// LS Electric XG5000 project: PLC MMI 2026 SCADA PLC 1
// PLC LSPLC
// module base 0 slot 0: Input/Output Module:XBC-DR64H (DC 24V Input, Relay Output, 64 Contacts)
// module base 0 slot 1: Cnet:XBL-C21A (Cnet Module(RS-232C))
// module base 0 slot 2: FEnet:XBL-EMTA (Ethernet Module, Electrical Master)

PROGRAM DataIndikatorProses (task: Scan Program)

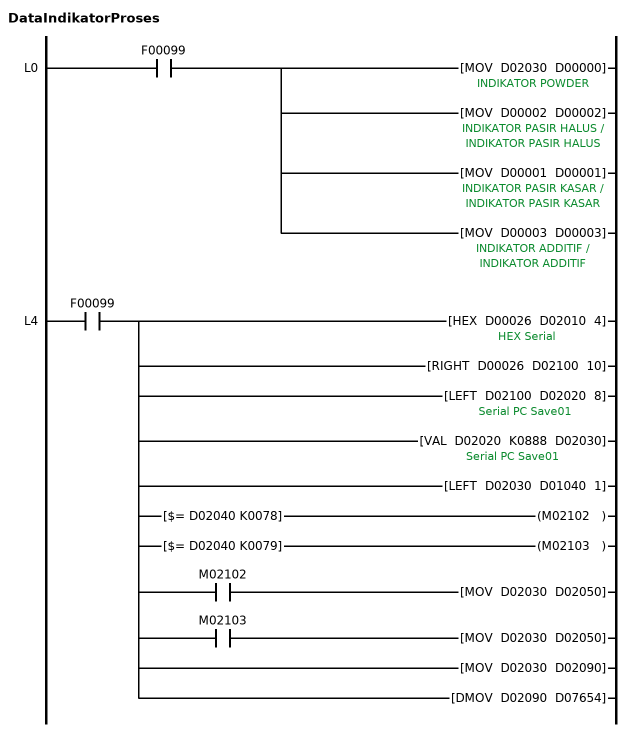
; L0
LOAD      F00099
MOV       D02030 D00000	// INDIKATOR POWDER
MOV       D00002 D00002	// INDIKATOR PASIR HALUS / INDIKATOR PASIR HALUS
MOV       D00001 D00001	// INDIKATOR PASIR KASAR / INDIKATOR PASIR KASAR
MOV       D00003 D00003	// INDIKATOR ADDITIF / INDIKATOR ADDITIF
; L4
LOAD      F00099
HEX       D00026 D02010 4	// HEX Serial
RIGHT     D00026 D02100 10
LEFT      D02100 D02020 8	// Serial PC Save01
VAL       D02020 K0888 D02030	// Serial PC Save01
LEFT      D02030 D01040 1
MPUSH
AND$=     D02040 K0078
OUT       M02102
MLOAD
AND$=     D02040 K0079
OUT       M02103
MLOAD
AND       M02102
MOV       D02030 D02050
MLOAD
AND       M02103
MOV       D02030 D02050
MPOP
MOV       D02030 D02090
DMOV      D02090 D07654

PROGRAM DataInverter (task: Scan Program)

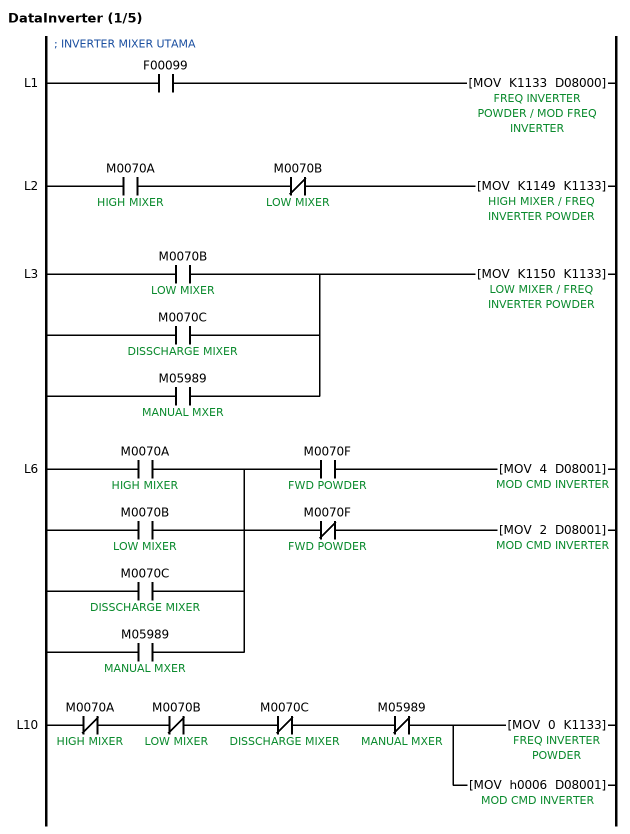
// INVERTER MIXER UTAMA
; L1
LOAD      F00099
MOV       K1133 D08000	// FREQ INVERTER POWDER / MOD FREQ INVERTER
; L2
LOAD      M0070A	// HIGH MIXER 
AND NOT   M0070B	// LOW MIXER 
MOV       K1149 K1133	// HIGH MIXER / FREQ INVERTER POWDER
; L3
LOAD      M0070B	// LOW MIXER 
OR        M0070C	// DISSCHARGE MIXER 
OR        M05989	// MANUAL MXER
MOV       K1150 K1133	// LOW MIXER / FREQ INVERTER POWDER
; L6
LOAD      M0070A	// HIGH MIXER 
OR        M0070B	// LOW MIXER 
OR        M0070C	// DISSCHARGE MIXER 
OR        M05989	// MANUAL MXER
MPUSH
AND       M0070F	// FWD POWDER
MOV       4 D08001	// MOD CMD INVERTER
MPOP
AND NOT   M0070F	// FWD POWDER
MOV       2 D08001	// MOD CMD INVERTER
; L10
LOAD NOT  M0070A	// HIGH MIXER 
AND NOT   M0070B	// LOW MIXER 
AND NOT   M0070C	// DISSCHARGE MIXER 
AND NOT   M05989	// MANUAL MXER
MOV       0 K1133	// FREQ INVERTER POWDER
MOV       h0006 D08001	// MOD CMD INVERTER

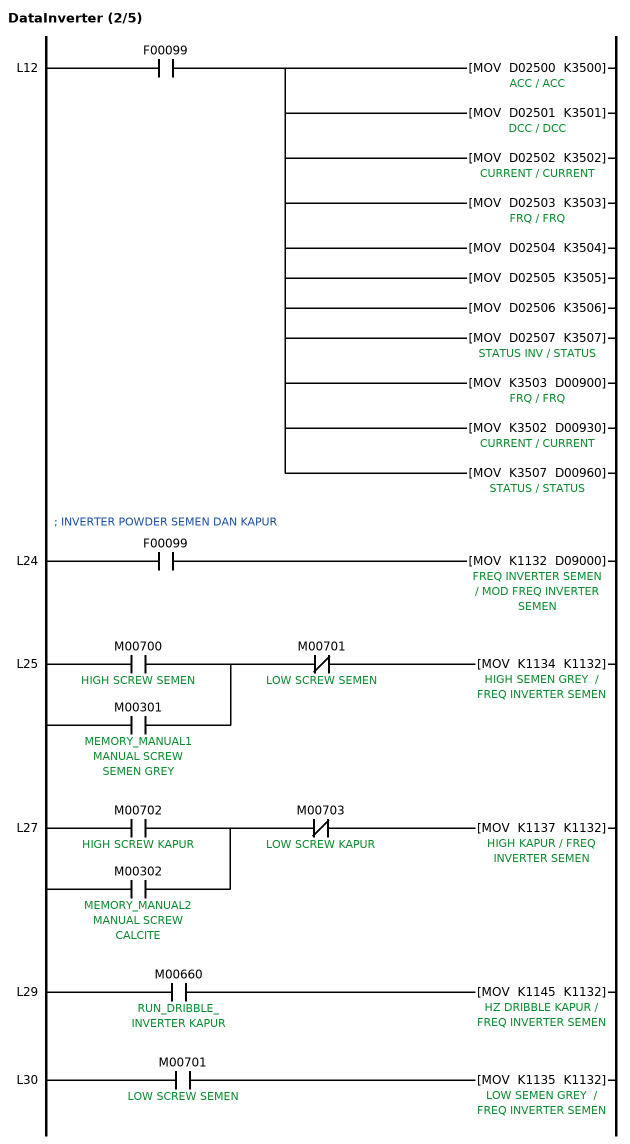
; L12
LOAD      F00099
MOV       D02500 K3500	// ACC / ACC
MOV       D02501 K3501	// DCC / DCC
MOV       D02502 K3502	// CURRENT / CURRENT
MOV       D02503 K3503	// FRQ / FRQ
MOV       D02504 K3504
MOV       D02505 K3505
MOV       D02506 K3506
MOV       D02507 K3507	// STATUS INV / STATUS
MOV       K3503 D00900	// FRQ / FRQ
MOV       K3502 D00930	// CURRENT / CURRENT
MOV       K3507 D00960	// STATUS / STATUS
// INVERTER POWDER SEMEN DAN KAPUR
; L24
LOAD      F00099
MOV       K1132 D09000	// FREQ INVERTER SEMEN  / MOD FREQ INVERTER SEMEN
; L25
LOAD      M00700	// HIGH SCREW SEMEN
OR        M00301	// MEMORY_MANUAL1 MANUAL SCREW SEMEN GREY 
AND NOT   M00701	// LOW SCREW SEMEN
MOV       K1134 K1132	// HIGH SEMEN GREY  / FREQ INVERTER SEMEN 
; L27
LOAD      M00702	// HIGH SCREW KAPUR
OR        M00302	// MEMORY_MANUAL2 MANUAL SCREW CALCITE
AND NOT   M00703	// LOW SCREW KAPUR
MOV       K1137 K1132	// HIGH KAPUR / FREQ INVERTER SEMEN 
; L29
LOAD      M00660	// RUN_DRIBBLE_INVERTER KAPUR
MOV       K1145 K1132	// HZ DRIBBLE KAPUR / FREQ INVERTER SEMEN 
; L30
LOAD      M00701	// LOW SCREW SEMEN
MOV       K1135 K1132	// LOW SEMEN GREY  / FREQ INVERTER SEMEN 

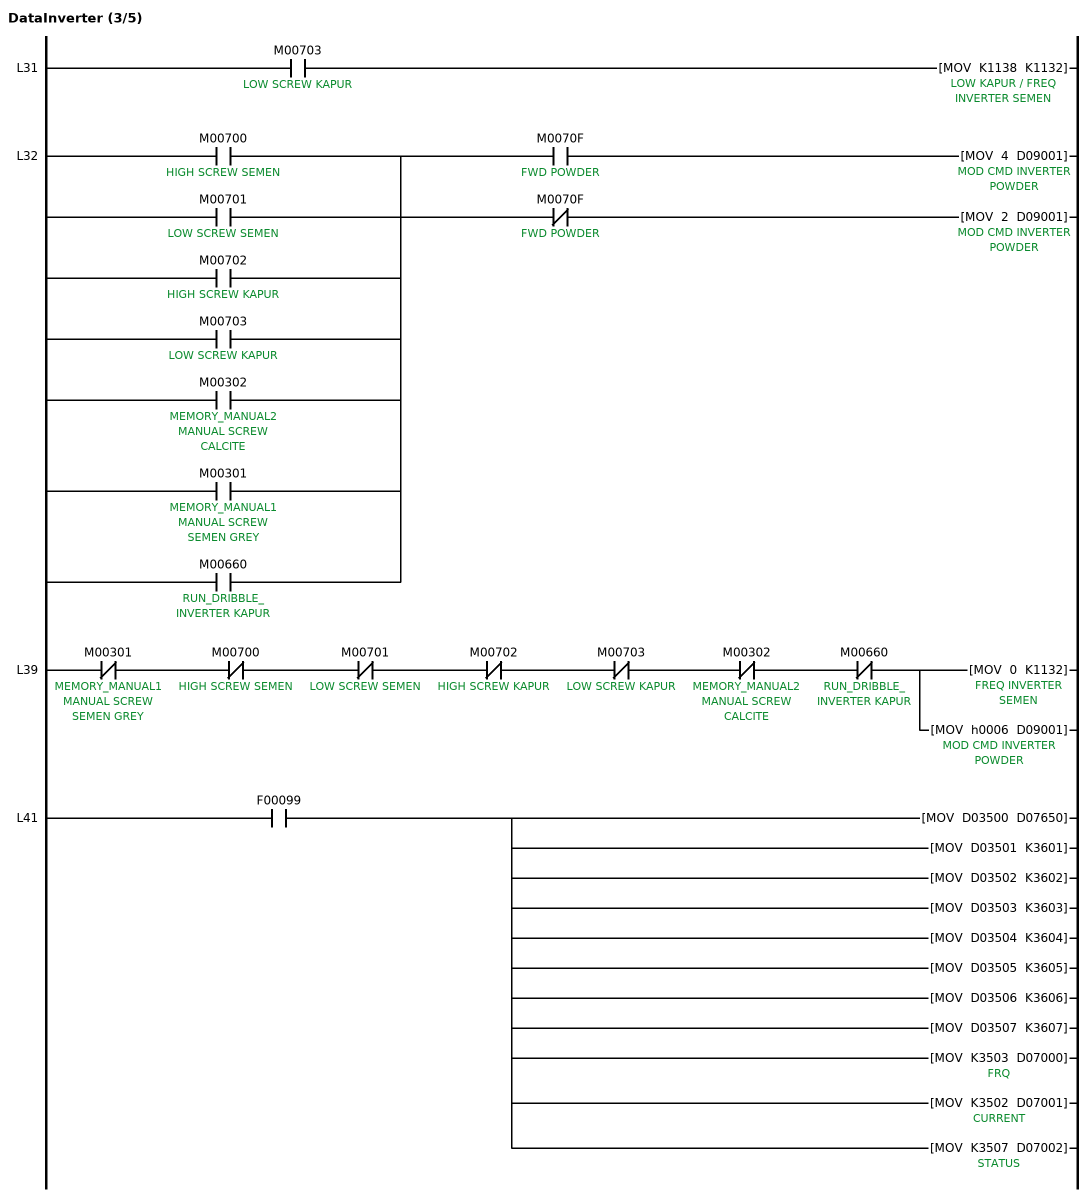
; L31
LOAD      M00703	// LOW SCREW KAPUR
MOV       K1138 K1132	// LOW KAPUR / FREQ INVERTER SEMEN 
; L32
LOAD      M00700	// HIGH SCREW SEMEN
OR        M00701	// LOW SCREW SEMEN
OR        M00702	// HIGH SCREW KAPUR
OR        M00703	// LOW SCREW KAPUR
OR        M00302	// MEMORY_MANUAL2 MANUAL SCREW CALCITE
OR        M00301	// MEMORY_MANUAL1 MANUAL SCREW SEMEN GREY 
OR        M00660	// RUN_DRIBBLE_INVERTER KAPUR
MPUSH
AND       M0070F	// FWD POWDER
MOV       4 D09001	// MOD CMD INVERTER POWDER
MPOP
AND NOT   M0070F	// FWD POWDER
MOV       2 D09001	// MOD CMD INVERTER POWDER
; L39
LOAD NOT  M00301	// MEMORY_MANUAL1 MANUAL SCREW SEMEN GREY 
AND NOT   M00700	// HIGH SCREW SEMEN
AND NOT   M00701	// LOW SCREW SEMEN
AND NOT   M00702	// HIGH SCREW KAPUR
AND NOT   M00703	// LOW SCREW KAPUR
AND NOT   M00302	// MEMORY_MANUAL2 MANUAL SCREW CALCITE
AND NOT   M00660	// RUN_DRIBBLE_INVERTER KAPUR
MOV       0 K1132	// FREQ INVERTER SEMEN 
MOV       h0006 D09001	// MOD CMD INVERTER POWDER
; L41
LOAD      F00099
MOV       D03500 D07650
MOV       D03501 K3601
MOV       D03502 K3602
MOV       D03503 K3603
MOV       D03504 K3604
MOV       D03505 K3605
MOV       D03506 K3606
MOV       D03507 K3607
MOV       K3503 D07000	// FRQ
MOV       K3502 D07001	// CURRENT
MOV       K3507 D07002	// STATUS

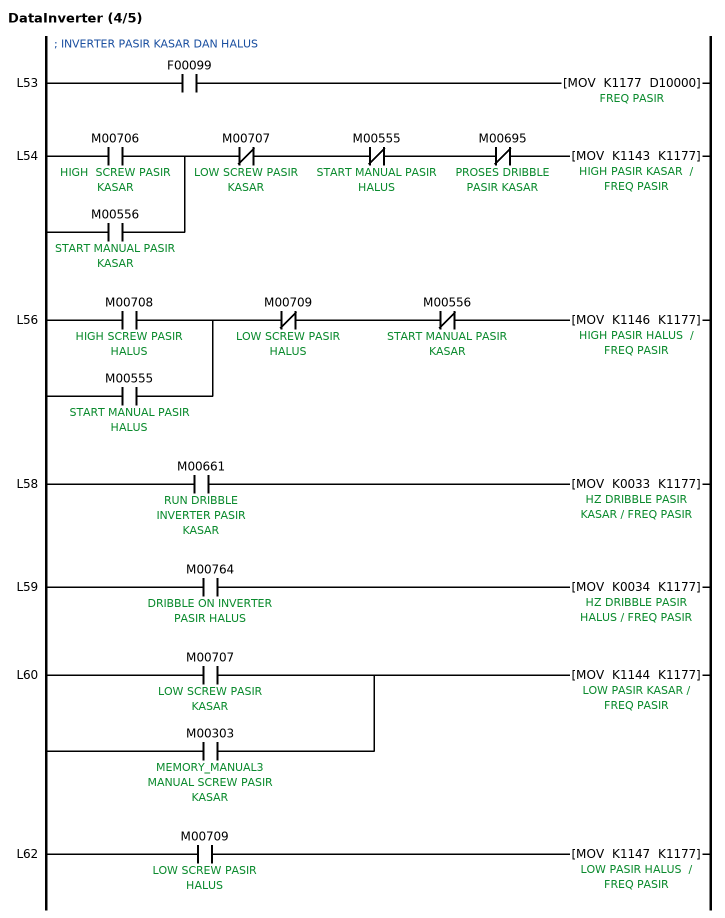
// INVERTER PASIR KASAR DAN HALUS
; L53
LOAD      F00099
MOV       K1177 D10000	// FREQ PASIR
; L54
LOAD      M00706	// HIGH  SCREW PASIR KASAR
OR        M00556	// START MANUAL PASIR KASAR
AND NOT   M00707	// LOW SCREW PASIR KASAR
AND NOT   M00555	// START MANUAL PASIR HALUS
AND NOT   M00695	// PROSES DRIBBLE PASIR KASAR
MOV       K1143 K1177	// HIGH PASIR KASAR  / FREQ PASIR
; L56
LOAD      M00708	// HIGH SCREW PASIR HALUS
OR        M00555	// START MANUAL PASIR HALUS
AND NOT   M00709	// LOW SCREW PASIR HALUS 
AND NOT   M00556	// START MANUAL PASIR KASAR
MOV       K1146 K1177	// HIGH PASIR HALUS  / FREQ PASIR
; L58
LOAD      M00661	// RUN DRIBBLE INVERTER PASIR KASAR
MOV       K0033 K1177	// HZ DRIBBLE PASIR KASAR / FREQ PASIR
; L59
LOAD      M00764	// DRIBBLE ON INVERTER PASIR HALUS
MOV       K0034 K1177	// HZ DRIBBLE PASIR HALUS / FREQ PASIR
; L60
LOAD      M00707	// LOW SCREW PASIR KASAR
OR        M00303	// MEMORY_MANUAL3 MANUAL SCREW PASIR KASAR
MOV       K1144 K1177	// LOW PASIR KASAR / FREQ PASIR
; L62
LOAD      M00709	// LOW SCREW PASIR HALUS 
MOV       K1147 K1177	// LOW PASIR HALUS  / FREQ PASIR

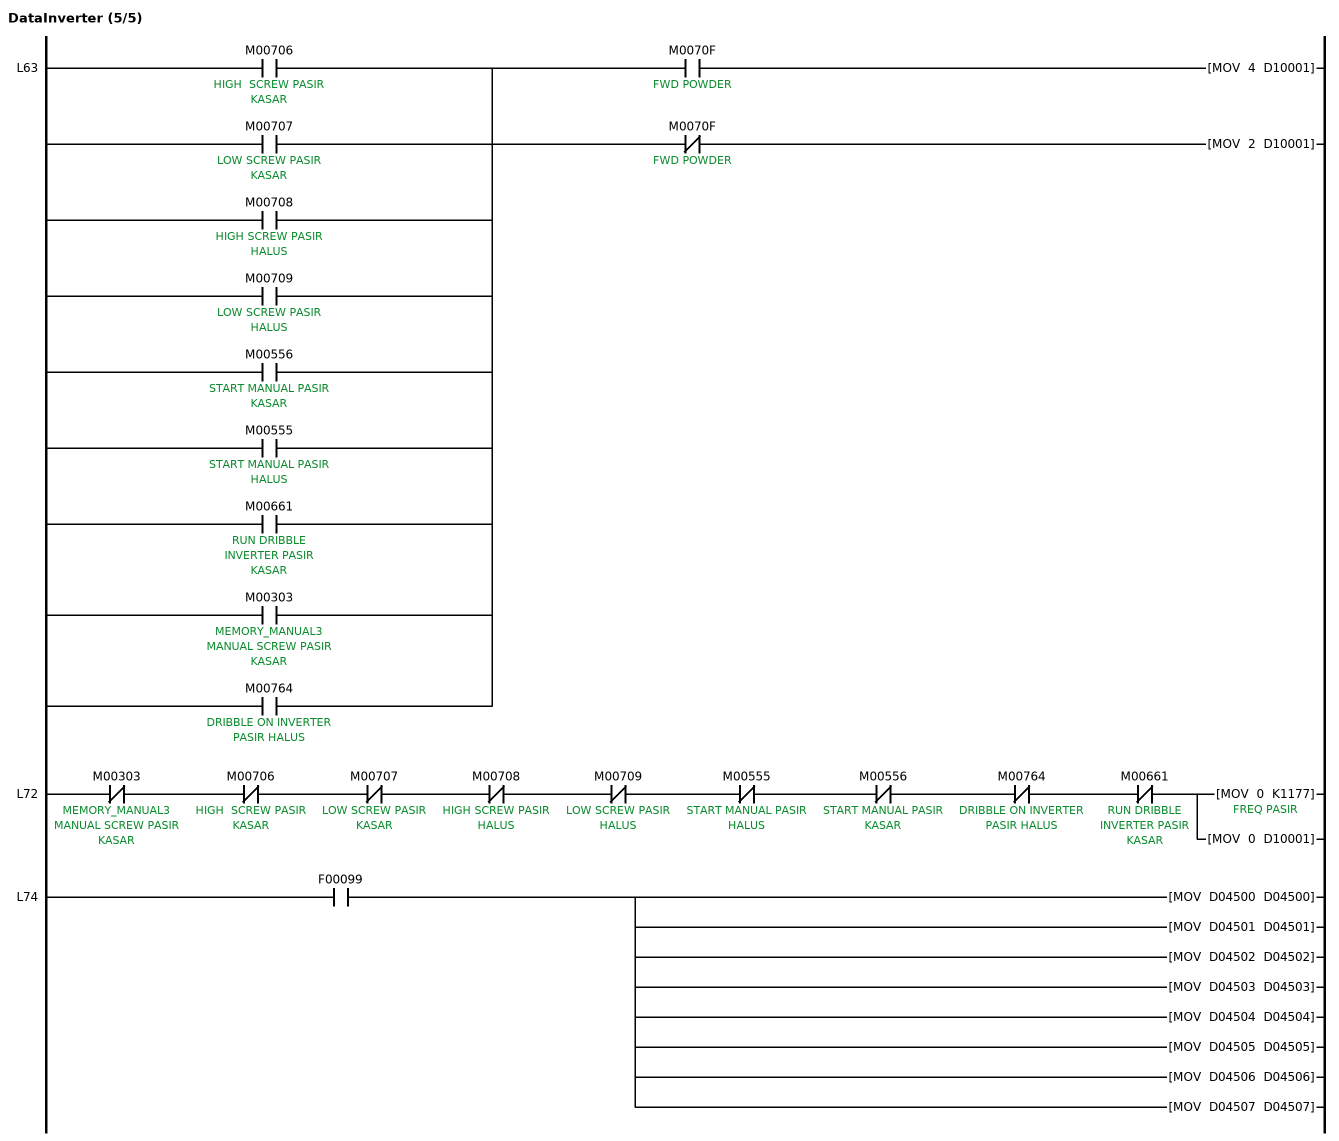
; L63
LOAD      M00706	// HIGH  SCREW PASIR KASAR
OR        M00707	// LOW SCREW PASIR KASAR
OR        M00708	// HIGH SCREW PASIR HALUS
OR        M00709	// LOW SCREW PASIR HALUS 
OR        M00556	// START MANUAL PASIR KASAR
OR        M00555	// START MANUAL PASIR HALUS
OR        M00661	// RUN DRIBBLE INVERTER PASIR KASAR
OR        M00303	// MEMORY_MANUAL3 MANUAL SCREW PASIR KASAR
OR        M00764	// DRIBBLE ON INVERTER PASIR HALUS
MPUSH
AND       M0070F	// FWD POWDER
MOV       4 D10001
MPOP
AND NOT   M0070F	// FWD POWDER
MOV       2 D10001
; L72
LOAD NOT  M00303	// MEMORY_MANUAL3 MANUAL SCREW PASIR KASAR
AND NOT   M00706	// HIGH  SCREW PASIR KASAR
AND NOT   M00707	// LOW SCREW PASIR KASAR
AND NOT   M00708	// HIGH SCREW PASIR HALUS
AND NOT   M00709	// LOW SCREW PASIR HALUS 
AND NOT   M00555	// START MANUAL PASIR HALUS
AND NOT   M00556	// START MANUAL PASIR KASAR
AND NOT   M00764	// DRIBBLE ON INVERTER PASIR HALUS
AND NOT   M00661	// RUN DRIBBLE INVERTER PASIR KASAR
MOV       0 K1177	// FREQ PASIR
MOV       0 D10001
; L74
LOAD      F00099
MOV       D04500 D04500
MOV       D04501 D04501
MOV       D04502 D04502
MOV       D04503 D04503
MOV       D04504 D04504
MOV       D04505 D04505
MOV       D04506 D04506
MOV       D04507 D04507

PROGRAM FormulaSet (task: Scan Program)

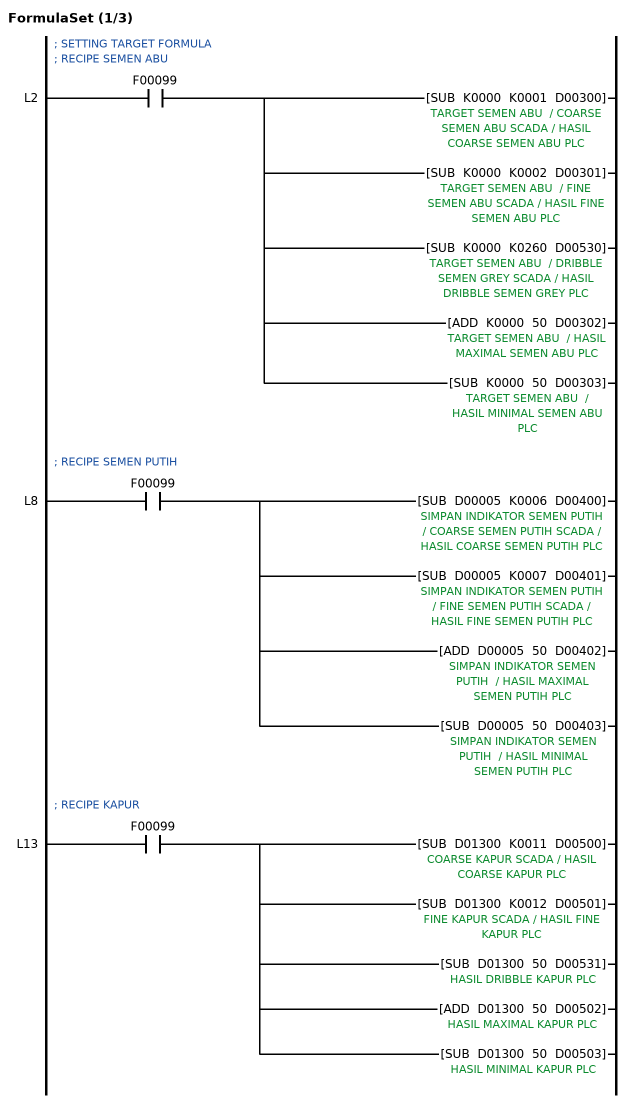
// SETTING TARGET FORMULA
// RECIPE SEMEN ABU
; L2
LOAD      F00099
SUB       K0000 K0001 D00300	// TARGET SEMEN ABU  / COARSE SEMEN ABU SCADA / HASIL COARSE SEMEN ABU PLC
SUB       K0000 K0002 D00301	// TARGET SEMEN ABU  / FINE SEMEN ABU SCADA / HASIL FINE SEMEN ABU PLC
SUB       K0000 K0260 D00530	// TARGET SEMEN ABU  / DRIBBLE SEMEN GREY SCADA / HASIL DRIBBLE SEMEN GREY PLC
ADD       K0000 50 D00302	// TARGET SEMEN ABU  / HASIL MAXIMAL SEMEN ABU PLC
SUB       K0000 50 D00303	// TARGET SEMEN ABU  / HASIL MINIMAL SEMEN ABU PLC
// RECIPE SEMEN PUTIH
; L8
LOAD      F00099
SUB       D00005 K0006 D00400	// SIMPAN INDIKATOR SEMEN PUTIH  / COARSE SEMEN PUTIH SCADA / HASIL COARSE SEMEN PUTIH PLC
SUB       D00005 K0007 D00401	// SIMPAN INDIKATOR SEMEN PUTIH  / FINE SEMEN PUTIH SCADA / HASIL FINE SEMEN PUTIH PLC 
ADD       D00005 50 D00402	// SIMPAN INDIKATOR SEMEN PUTIH  / HASIL MAXIMAL SEMEN PUTIH PLC 
SUB       D00005 50 D00403	// SIMPAN INDIKATOR SEMEN PUTIH  / HASIL MINIMAL SEMEN PUTIH PLC
// RECIPE KAPUR
; L13
LOAD      F00099
SUB       D01300 K0011 D00500	// COARSE KAPUR SCADA / HASIL COARSE KAPUR PLC
SUB       D01300 K0012 D00501	// FINE KAPUR SCADA / HASIL FINE KAPUR PLC 
SUB       D01300 50 D00531	// HASIL DRIBBLE KAPUR PLC 
ADD       D01300 50 D00502	// HASIL MAXIMAL KAPUR PLC 
SUB       D01300 50 D00503	// HASIL MINIMAL KAPUR PLC 

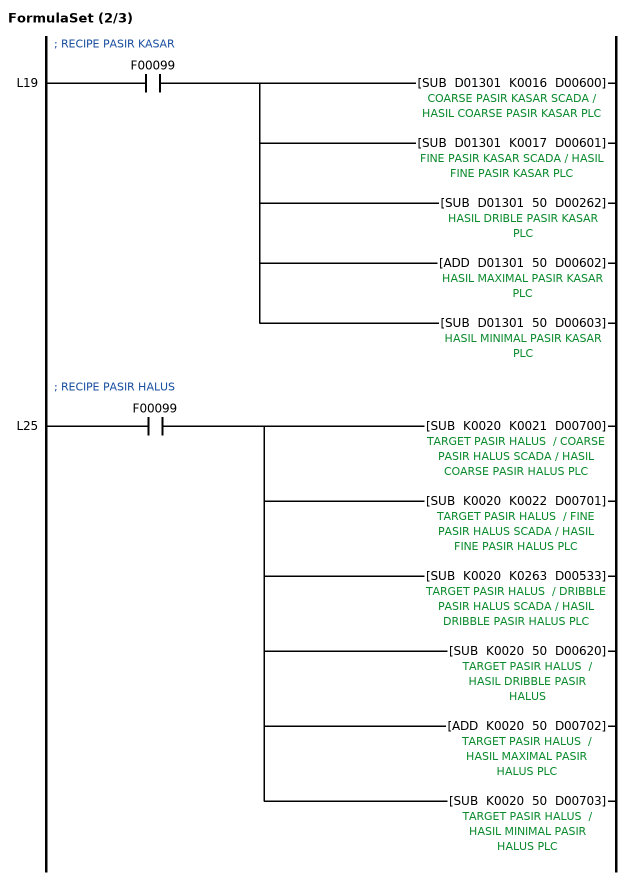
// RECIPE PASIR KASAR
; L19
LOAD      F00099
SUB       D01301 K0016 D00600	// COARSE PASIR KASAR SCADA / HASIL COARSE PASIR KASAR PLC
SUB       D01301 K0017 D00601	// FINE PASIR KASAR SCADA / HASIL FINE PASIR KASAR PLC
SUB       D01301 50 D00262	// HASIL DRIBLE PASIR KASAR PLC
ADD       D01301 50 D00602	// HASIL MAXIMAL PASIR KASAR PLC
SUB       D01301 50 D00603	// HASIL MINIMAL PASIR KASAR PLC
// RECIPE PASIR HALUS
; L25
LOAD      F00099
SUB       K0020 K0021 D00700	// TARGET PASIR HALUS  / COARSE PASIR HALUS SCADA / HASIL COARSE PASIR HALUS PLC
SUB       K0020 K0022 D00701	// TARGET PASIR HALUS  / FINE PASIR HALUS SCADA / HASIL FINE PASIR HALUS PLC
SUB       K0020 K0263 D00533	// TARGET PASIR HALUS  / DRIBBLE PASIR HALUS SCADA / HASIL DRIBBLE PASIR HALUS PLC
SUB       K0020 50 D00620	// TARGET PASIR HALUS  / HASIL DRIBBLE PASIR HALUS
ADD       K0020 50 D00702	// TARGET PASIR HALUS  / HASIL MAXIMAL PASIR HALUS PLC
SUB       K0020 50 D00703	// TARGET PASIR HALUS  / HASIL MINIMAL PASIR HALUS PLC

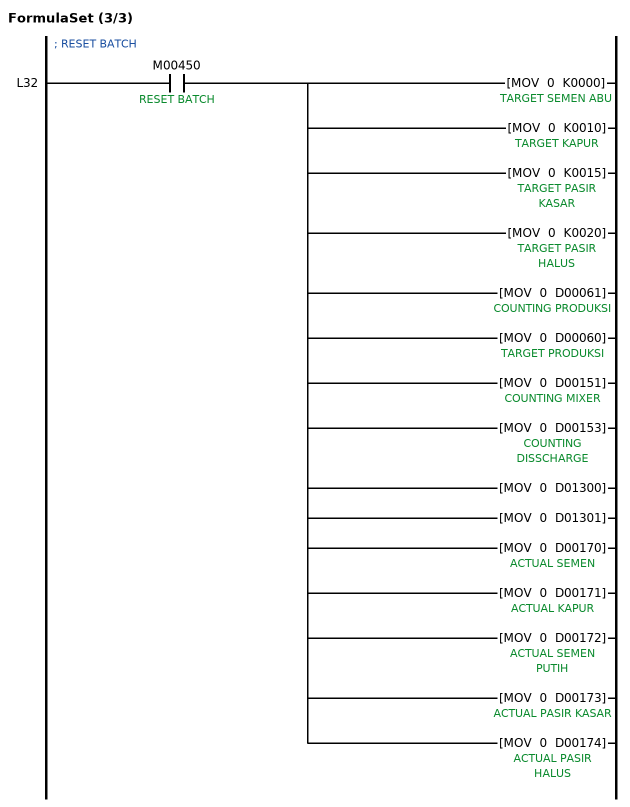
// RESET BATCH
; L32
LOAD      M00450	// RESET BATCH
MOV       0 K0000	// TARGET SEMEN ABU 
MOV       0 K0010	// TARGET KAPUR 
MOV       0 K0015	// TARGET PASIR KASAR
MOV       0 K0020	// TARGET PASIR HALUS 
MOV       0 D00061	// COUNTING PRODUKSI
MOV       0 D00060	// TARGET PRODUKSI
MOV       0 D00151	// COUNTING MIXER
MOV       0 D00153	// COUNTING DISSCHARGE
MOV       0 D01300
MOV       0 D01301
MOV       0 D00170	// ACTUAL SEMEN
MOV       0 D00171	// ACTUAL KAPUR
MOV       0 D00172	// ACTUAL SEMEN PUTIH
MOV       0 D00173	// ACTUAL PASIR KASAR
MOV       0 D00174	// ACTUAL PASIR HALUS

PROGRAM DigitalInput (task: Scan Program)

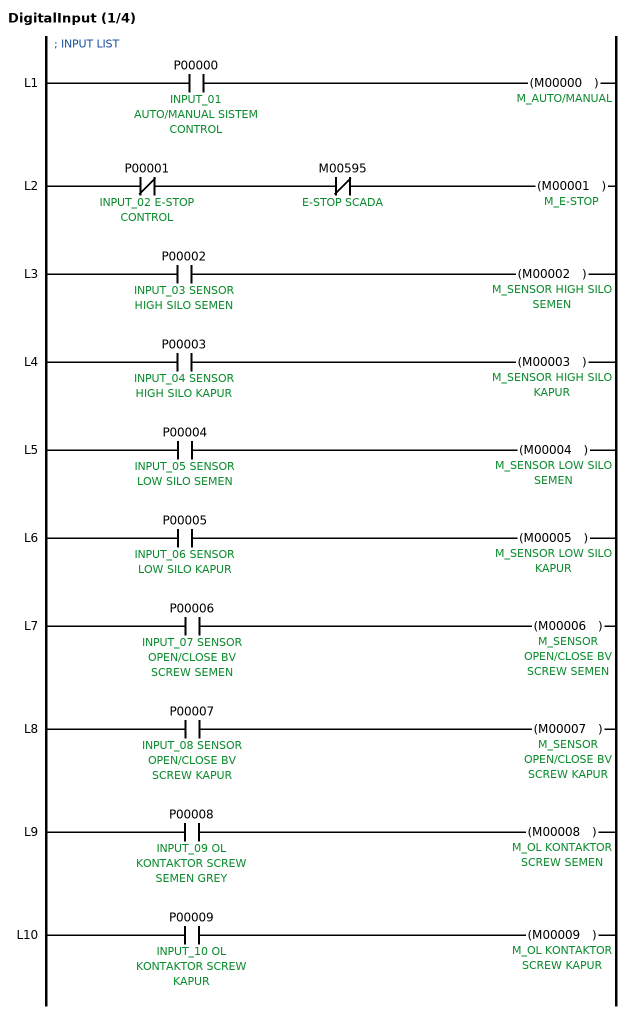
// INPUT LIST
; L1
LOAD      P00000	// INPUT_01 AUTO/MANUAL SISTEM CONTROL
OUT       M00000	// M_AUTO/MANUAL
; L2
LOAD NOT  P00001	// INPUT_02 E-STOP CONTROL 
AND NOT   M00595	// E-STOP SCADA
OUT       M00001	// M_E-STOP
; L3
LOAD      P00002	// INPUT_03 SENSOR HIGH SILO SEMEN
OUT       M00002	// M_SENSOR HIGH SILO SEMEN 
; L4
LOAD      P00003	// INPUT_04 SENSOR HIGH SILO KAPUR
OUT       M00003	// M_SENSOR HIGH SILO KAPUR
; L5
LOAD      P00004	// INPUT_05 SENSOR LOW SILO SEMEN
OUT       M00004	// M_SENSOR LOW SILO SEMEN 
; L6
LOAD      P00005	// INPUT_06 SENSOR LOW SILO KAPUR
OUT       M00005	// M_SENSOR LOW SILO KAPUR
; L7
LOAD      P00006	// INPUT_07 SENSOR OPEN/CLOSE BV SCREW SEMEN
OUT       M00006	// M_SENSOR OPEN/CLOSE BV SCREW SEMEN
; L8
LOAD      P00007	// INPUT_08 SENSOR OPEN/CLOSE BV SCREW KAPUR
OUT       M00007	// M_SENSOR OPEN/CLOSE BV SCREW KAPUR
; L9
LOAD      P00008	// INPUT_09 OL KONTAKTOR SCREW SEMEN GREY 
OUT       M00008	// M_OL KONTAKTOR SCREW SEMEN
; L10
LOAD      P00009	// INPUT_10 OL KONTAKTOR SCREW KAPUR
OUT       M00009	// M_OL KONTAKTOR SCREW KAPUR

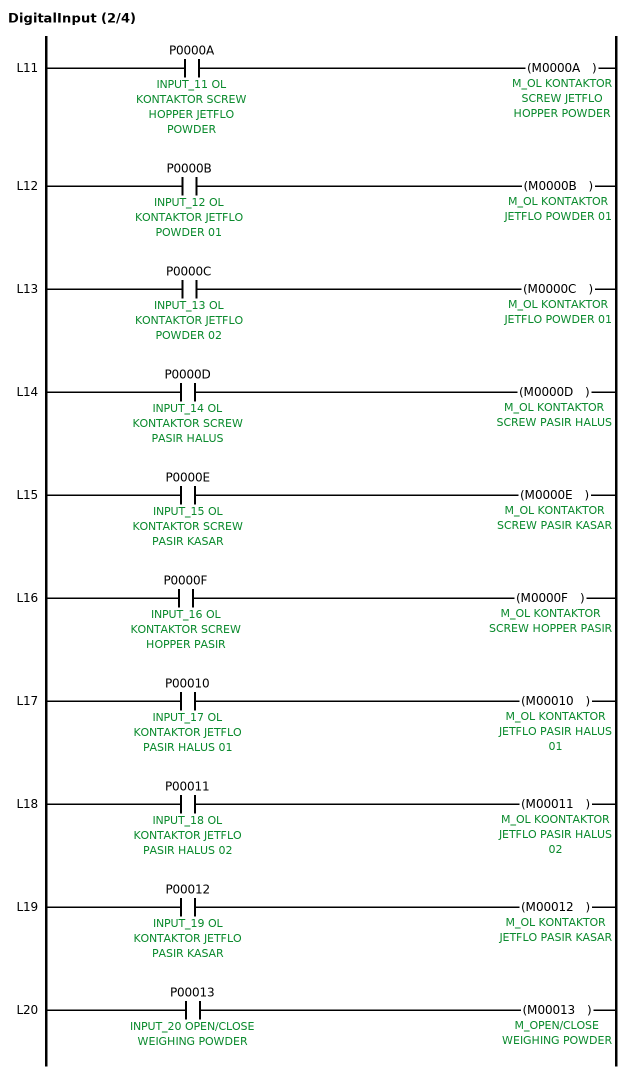
; L11
LOAD      P0000A	// INPUT_11 OL KONTAKTOR SCREW HOPPER JETFLO POWDER
OUT       M0000A	// M_OL KONTAKTOR SCREW JETFLO HOPPER POWDER
; L12
LOAD      P0000B	// INPUT_12 OL KONTAKTOR JETFLO POWDER 01
OUT       M0000B	// M_OL KONTAKTOR JETFLO POWDER 01
; L13
LOAD      P0000C	// INPUT_13 OL KONTAKTOR JETFLO POWDER 02
OUT       M0000C	// M_OL KONTAKTOR JETFLO POWDER 01
; L14
LOAD      P0000D	// INPUT_14 OL KONTAKTOR SCREW PASIR HALUS 
OUT       M0000D	// M_OL KONTAKTOR SCREW PASIR HALUS 
; L15
LOAD      P0000E	// INPUT_15 OL KONTAKTOR SCREW PASIR KASAR
OUT       M0000E	// M_OL KONTAKTOR SCREW PASIR KASAR
; L16
LOAD      P0000F	// INPUT_16 OL KONTAKTOR SCREW HOPPER PASIR 
OUT       M0000F	// M_OL KONTAKTOR SCREW HOPPER PASIR
; L17
LOAD      P00010	// INPUT_17 OL KONTAKTOR JETFLO PASIR HALUS 01
OUT       M00010	// M_OL KONTAKTOR JETFLO PASIR HALUS 01
; L18
LOAD      P00011	// INPUT_18 OL KONTAKTOR JETFLO PASIR HALUS 02
OUT       M00011	// M_OL KOONTAKTOR JETFLO PASIR HALUS 02
; L19
LOAD      P00012	// INPUT_19 OL KONTAKTOR JETFLO PASIR KASAR 
OUT       M00012	// M_OL KONTAKTOR JETFLO PASIR KASAR
; L20
LOAD      P00013	// INPUT_20 OPEN/CLOSE WEIGHING POWDER
OUT       M00013	// M_OPEN/CLOSE WEIGHING POWDER

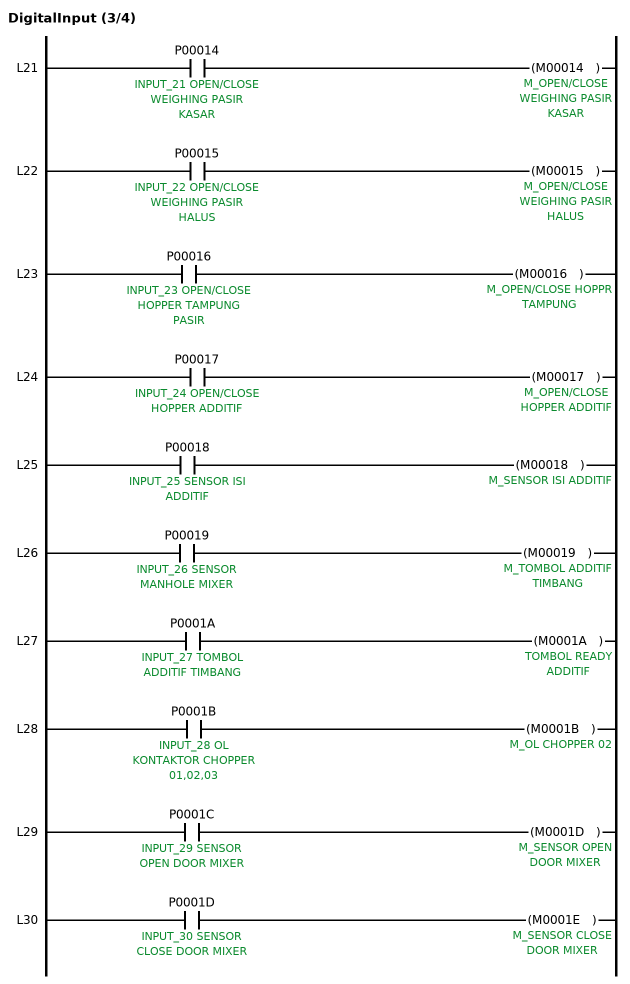
; L21
LOAD      P00014	// INPUT_21 OPEN/CLOSE WEIGHING PASIR KASAR
OUT       M00014	// M_OPEN/CLOSE WEIGHING PASIR KASAR
; L22
LOAD      P00015	// INPUT_22 OPEN/CLOSE WEIGHING PASIR HALUS
OUT       M00015	// M_OPEN/CLOSE WEIGHING PASIR HALUS 
; L23
LOAD      P00016	// INPUT_23 OPEN/CLOSE HOPPER TAMPUNG PASIR
OUT       M00016	// M_OPEN/CLOSE HOPPR TAMPUNG
; L24
LOAD      P00017	// INPUT_24 OPEN/CLOSE HOPPER ADDITIF
OUT       M00017	// M_OPEN/CLOSE HOPPER ADDITIF
; L25
LOAD      P00018	// INPUT_25 SENSOR ISI ADDITIF
OUT       M00018	// M_SENSOR ISI ADDITIF
; L26
LOAD      P00019	// INPUT_26 SENSOR MANHOLE MIXER
OUT       M00019	// M_TOMBOL ADDITIF TIMBANG
; L27
LOAD      P0001A	// INPUT_27 TOMBOL ADDITIF TIMBANG 
OUT       M0001A	// TOMBOL READY ADDITIF
; L28
LOAD      P0001B	// INPUT_28 OL KONTAKTOR CHOPPER 01,02,03
OUT       M0001B	// M_OL CHOPPER 02
; L29
LOAD      P0001C	// INPUT_29 SENSOR OPEN DOOR MIXER
OUT       M0001D	// M_SENSOR OPEN DOOR MIXER 
; L30
LOAD      P0001D	// INPUT_30 SENSOR CLOSE DOOR MIXER
OUT       M0001E	// M_SENSOR CLOSE DOOR MIXER

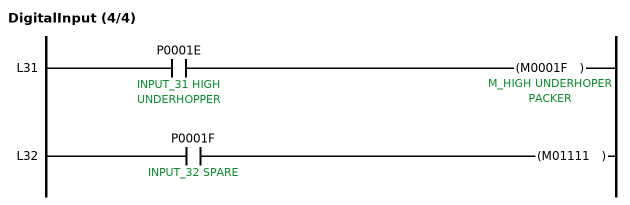
; L31
LOAD      P0001E	// INPUT_31 HIGH UNDERHOPPER
OUT       M0001F	// M_HIGH UNDERHOPER PACKER
; L32
LOAD      P0001F	// INPUT_32 SPARE
OUT       M01111

PROGRAM DigitalOutput (task: Scan Program)

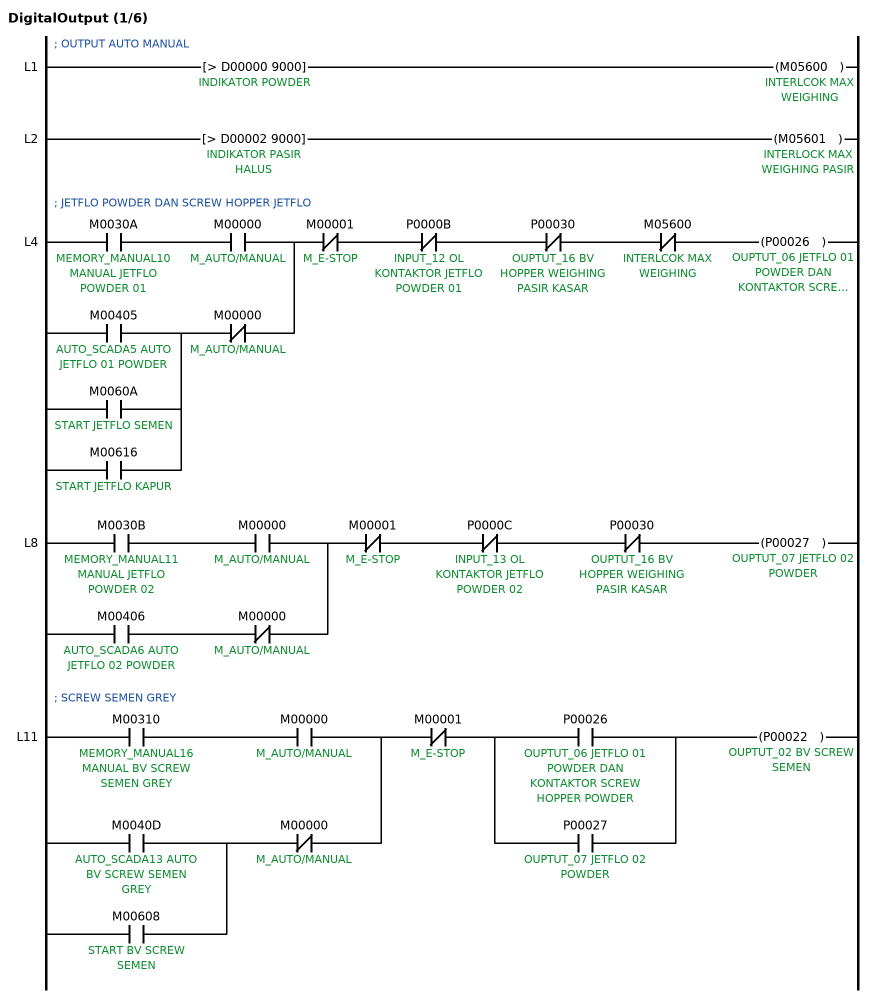
// OUTPUT AUTO MANUAL
; L1
LOAD>     D00000 9000	// INDIKATOR POWDER
OUT       M05600	// INTERLCOK MAX WEIGHING
; L2
LOAD>     D00002 9000	// INDIKATOR PASIR HALUS
OUT       M05601	// INTERLOCK MAX WEIGHING PASIR
// JETFLO POWDER DAN SCREW HOPPER JETFLO
; L4
LOAD      M0030A	// MEMORY_MANUAL10 MANUAL JETFLO POWDER 01 
AND       M00000	// M_AUTO/MANUAL
LOAD      M00405	// AUTO_SCADA5 AUTO JETFLO 01 POWDER
OR        M0060A	// START JETFLO SEMEN
OR        M00616	// START JETFLO KAPUR
AND NOT   M00000	// M_AUTO/MANUAL
OR LOAD
AND NOT   M00001	// M_E-STOP
AND NOT   P0000B	// INPUT_12 OL KONTAKTOR JETFLO POWDER 01
AND NOT   P00030	// OUPTUT_16 BV HOPPER WEIGHING PASIR KASAR
AND NOT   M05600	// INTERLCOK MAX WEIGHING
OUT       P00026	// OUPTUT_06 JETFLO 01 POWDER DAN KONTAKTOR SCREW HOPPER POWDER
; L8
LOAD      M0030B	// MEMORY_MANUAL11 MANUAL JETFLO POWDER 02 
AND       M00000	// M_AUTO/MANUAL
LOAD      M00406	// AUTO_SCADA6 AUTO JETFLO 02 POWDER
AND NOT   M00000	// M_AUTO/MANUAL
OR LOAD
AND NOT   M00001	// M_E-STOP
AND NOT   P0000C	// INPUT_13 OL KONTAKTOR JETFLO POWDER 02
AND NOT   P00030	// OUPTUT_16 BV HOPPER WEIGHING PASIR KASAR
OUT       P00027	// OUPTUT_07 JETFLO 02 POWDER 
// SCREW SEMEN GREY
; L11
LOAD      M00310	// MEMORY_MANUAL16 MANUAL BV SCREW SEMEN GREY 
AND       M00000	// M_AUTO/MANUAL
LOAD      M0040D	// AUTO_SCADA13 AUTO BV SCREW SEMEN GREY 
OR        M00608	// START BV SCREW SEMEN 
AND NOT   M00000	// M_AUTO/MANUAL
OR LOAD
AND NOT   M00001	// M_E-STOP
LOAD      P00026	// OUPTUT_06 JETFLO 01 POWDER DAN KONTAKTOR SCREW HOPPER POWDER
OR        P00027	// OUPTUT_07 JETFLO 02 POWDER 
AND LOAD
OUT       P00022	// OUPTUT_02 BV SCREW SEMEN

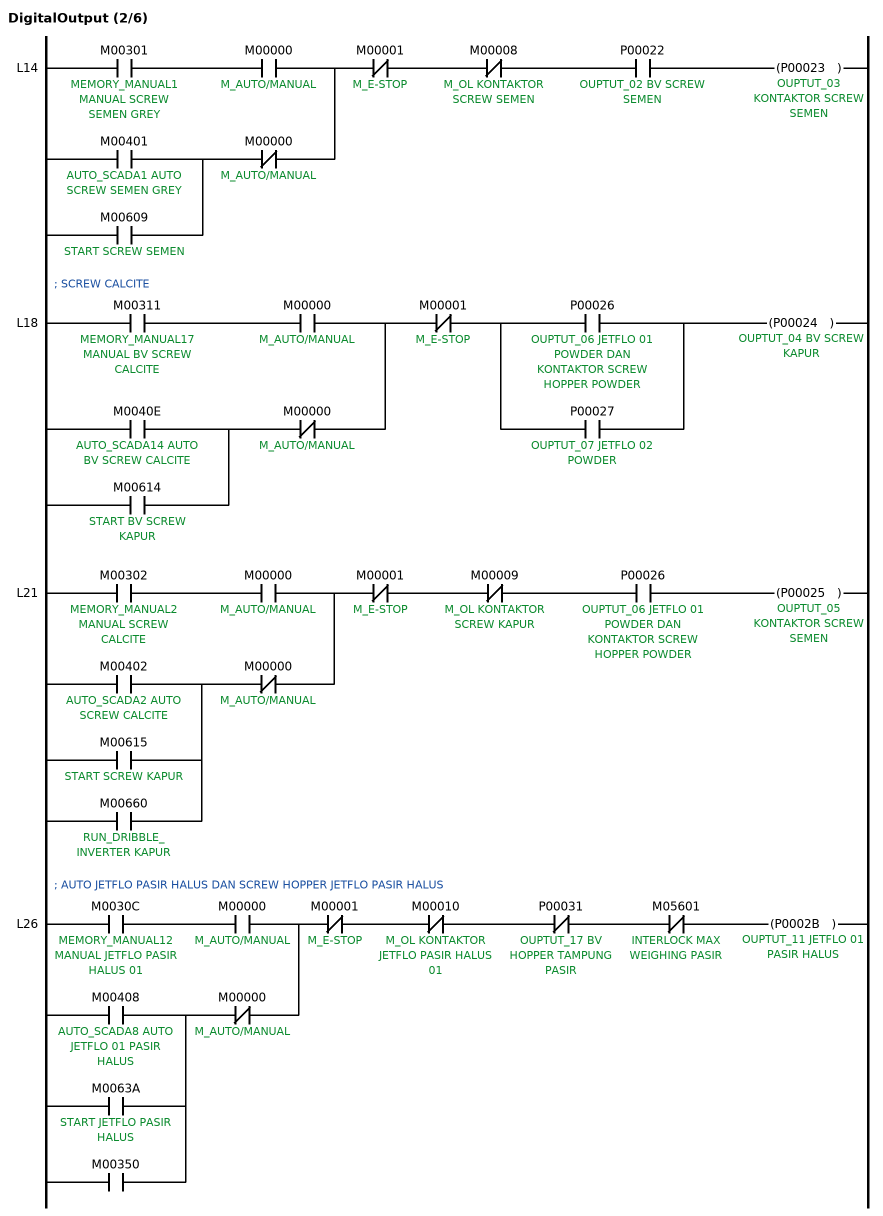
; L14
LOAD      M00301	// MEMORY_MANUAL1 MANUAL SCREW SEMEN GREY 
AND       M00000	// M_AUTO/MANUAL
LOAD      M00401	// AUTO_SCADA1 AUTO SCREW SEMEN GREY 
OR        M00609	// START SCREW SEMEN
AND NOT   M00000	// M_AUTO/MANUAL
OR LOAD
AND NOT   M00001	// M_E-STOP
AND NOT   M00008	// M_OL KONTAKTOR SCREW SEMEN
AND       P00022	// OUPTUT_02 BV SCREW SEMEN
OUT       P00023	// OUPTUT_03 KONTAKTOR SCREW SEMEN
// SCREW CALCITE
; L18
LOAD      M00311	// MEMORY_MANUAL17 MANUAL BV SCREW CALCITE
AND       M00000	// M_AUTO/MANUAL
LOAD      M0040E	// AUTO_SCADA14 AUTO BV SCREW CALCITE
OR        M00614	// START BV SCREW KAPUR
AND NOT   M00000	// M_AUTO/MANUAL
OR LOAD
AND NOT   M00001	// M_E-STOP
LOAD      P00026	// OUPTUT_06 JETFLO 01 POWDER DAN KONTAKTOR SCREW HOPPER POWDER
OR        P00027	// OUPTUT_07 JETFLO 02 POWDER 
AND LOAD
OUT       P00024	// OUPTUT_04 BV SCREW KAPUR
; L21
LOAD      M00302	// MEMORY_MANUAL2 MANUAL SCREW CALCITE
AND       M00000	// M_AUTO/MANUAL
LOAD      M00402	// AUTO_SCADA2 AUTO SCREW CALCITE
OR        M00615	// START SCREW KAPUR
OR        M00660	// RUN_DRIBBLE_INVERTER KAPUR
AND NOT   M00000	// M_AUTO/MANUAL
OR LOAD
AND NOT   M00001	// M_E-STOP
AND NOT   M00009	// M_OL KONTAKTOR SCREW KAPUR
AND       P00026	// OUPTUT_06 JETFLO 01 POWDER DAN KONTAKTOR SCREW HOPPER POWDER
OUT       P00025	// OUPTUT_05 KONTAKTOR SCREW SEMEN
// AUTO JETFLO PASIR HALUS DAN SCREW HOPPER JETFLO PASIR HALUS
; L26
LOAD      M0030C	// MEMORY_MANUAL12 MANUAL JETFLO PASIR HALUS 01 
AND       M00000	// M_AUTO/MANUAL
LOAD      M00408	// AUTO_SCADA8 AUTO JETFLO 01 PASIR HALUS 
OR        M0063A	// START JETFLO PASIR  HALUS
OR        M00350
AND NOT   M00000	// M_AUTO/MANUAL
OR LOAD
AND NOT   M00001	// M_E-STOP
AND NOT   M00010	// M_OL KONTAKTOR JETFLO PASIR HALUS 01
AND NOT   P00031	// OUPTUT_17 BV HOPPER TAMPUNG PASIR
AND NOT   M05601	// INTERLOCK MAX WEIGHING PASIR
OUT       P0002B	// OUPTUT_11 JETFLO 01 PASIR HALUS

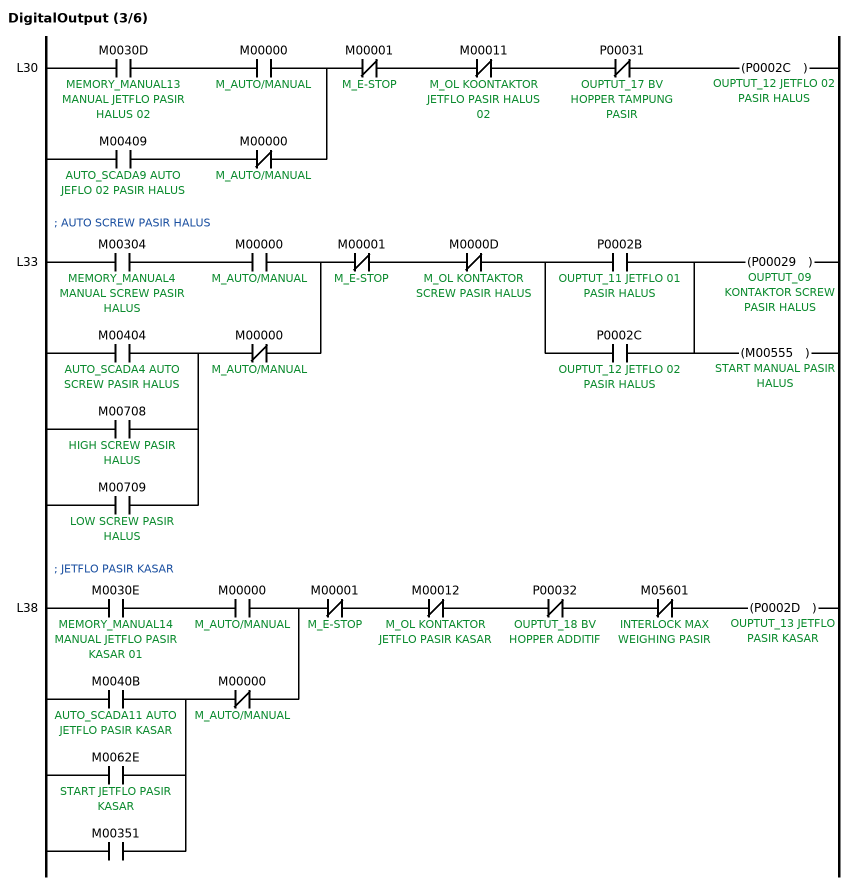
; L30
LOAD      M0030D	// MEMORY_MANUAL13 MANUAL JETFLO PASIR HALUS 02 
AND       M00000	// M_AUTO/MANUAL
LOAD      M00409	// AUTO_SCADA9 AUTO JEFLO 02 PASIR HALUS 
AND NOT   M00000	// M_AUTO/MANUAL
OR LOAD
AND NOT   M00001	// M_E-STOP
AND NOT   M00011	// M_OL KOONTAKTOR JETFLO PASIR HALUS 02
AND NOT   P00031	// OUPTUT_17 BV HOPPER TAMPUNG PASIR
OUT       P0002C	// OUPTUT_12 JETFLO 02 PASIR HALUS
// AUTO SCREW PASIR HALUS
; L33
LOAD      M00304	// MEMORY_MANUAL4 MANUAL SCREW PASIR HALUS 
AND       M00000	// M_AUTO/MANUAL
LOAD      M00404	// AUTO_SCADA4 AUTO SCREW PASIR HALUS 
OR        M00708	// HIGH SCREW PASIR HALUS
OR        M00709	// LOW SCREW PASIR HALUS 
AND NOT   M00000	// M_AUTO/MANUAL
OR LOAD
AND NOT   M00001	// M_E-STOP
AND NOT   M0000D	// M_OL KONTAKTOR SCREW PASIR HALUS 
LOAD      P0002B	// OUPTUT_11 JETFLO 01 PASIR HALUS
OR        P0002C	// OUPTUT_12 JETFLO 02 PASIR HALUS
AND LOAD
OUT       P00029	// OUPTUT_09 KONTAKTOR SCREW PASIR HALUS
OUT       M00555	// START MANUAL PASIR HALUS
// JETFLO PASIR KASAR
; L38
LOAD      M0030E	// MEMORY_MANUAL14 MANUAL JETFLO PASIR KASAR 01
AND       M00000	// M_AUTO/MANUAL
LOAD      M0040B	// AUTO_SCADA11 AUTO JETFLO PASIR KASAR 
OR        M0062E	// START JETFLO PASIR KASAR
OR        M00351
AND NOT   M00000	// M_AUTO/MANUAL
OR LOAD
AND NOT   M00001	// M_E-STOP
AND NOT   M00012	// M_OL KONTAKTOR JETFLO PASIR KASAR
AND NOT   P00032	// OUPTUT_18 BV HOPPER ADDITIF
AND NOT   M05601	// INTERLOCK MAX WEIGHING PASIR
OUT       P0002D	// OUPTUT_13 JETFLO PASIR KASAR

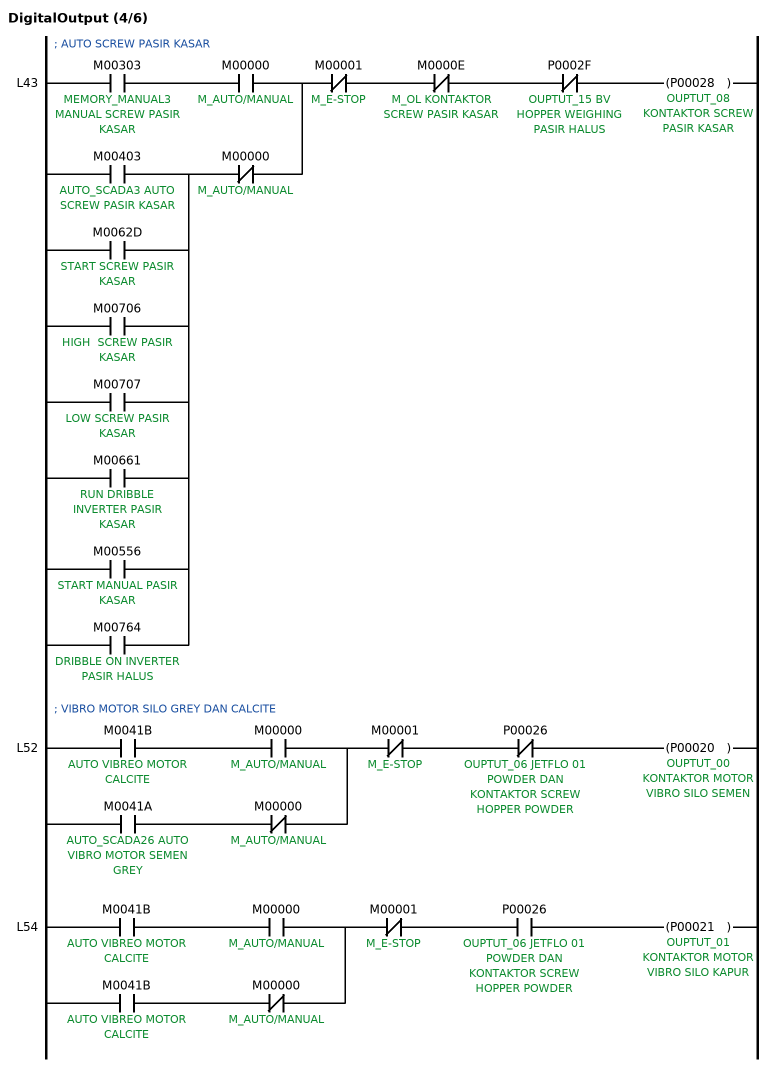
// AUTO SCREW PASIR KASAR
; L43
LOAD      M00303	// MEMORY_MANUAL3 MANUAL SCREW PASIR KASAR
AND       M00000	// M_AUTO/MANUAL
LOAD      M00403	// AUTO_SCADA3 AUTO SCREW PASIR KASAR 
OR        M0062D	// START SCREW PASIR KASAR
OR        M00706	// HIGH  SCREW PASIR KASAR
OR        M00707	// LOW SCREW PASIR KASAR
OR        M00661	// RUN DRIBBLE INVERTER PASIR KASAR
OR        M00556	// START MANUAL PASIR KASAR
OR        M00764	// DRIBBLE ON INVERTER PASIR HALUS
AND NOT   M00000	// M_AUTO/MANUAL
OR LOAD
AND NOT   M00001	// M_E-STOP
AND NOT   M0000E	// M_OL KONTAKTOR SCREW PASIR KASAR
AND NOT   P0002F	// OUPTUT_15 BV HOPPER WEIGHING PASIR HALUS
OUT       P00028	// OUPTUT_08 KONTAKTOR SCREW PASIR KASAR
// VIBRO MOTOR SILO GREY DAN CALCITE
; L52
LOAD      M0041B	// AUTO VIBREO MOTOR CALCITE
AND       M00000	// M_AUTO/MANUAL
LOAD      M0041A	// AUTO_SCADA26 AUTO VIBRO MOTOR SEMEN GREY 
AND NOT   M00000	// M_AUTO/MANUAL
OR LOAD
AND NOT   M00001	// M_E-STOP
AND NOT   P00026	// OUPTUT_06 JETFLO 01 POWDER DAN KONTAKTOR SCREW HOPPER POWDER
OUT       P00020	// OUPTUT_00 KONTAKTOR MOTOR VIBRO SILO SEMEN
; L54
LOAD      M0041B	// AUTO VIBREO MOTOR CALCITE
AND       M00000	// M_AUTO/MANUAL
LOAD      M0041B	// AUTO VIBREO MOTOR CALCITE
AND NOT   M00000	// M_AUTO/MANUAL
OR LOAD
AND NOT   M00001	// M_E-STOP
AND       P00026	// OUPTUT_06 JETFLO 01 POWDER DAN KONTAKTOR SCREW HOPPER POWDER
OUT       P00021	// OUPTUT_01 KONTAKTOR MOTOR VIBRO SILO KAPUR

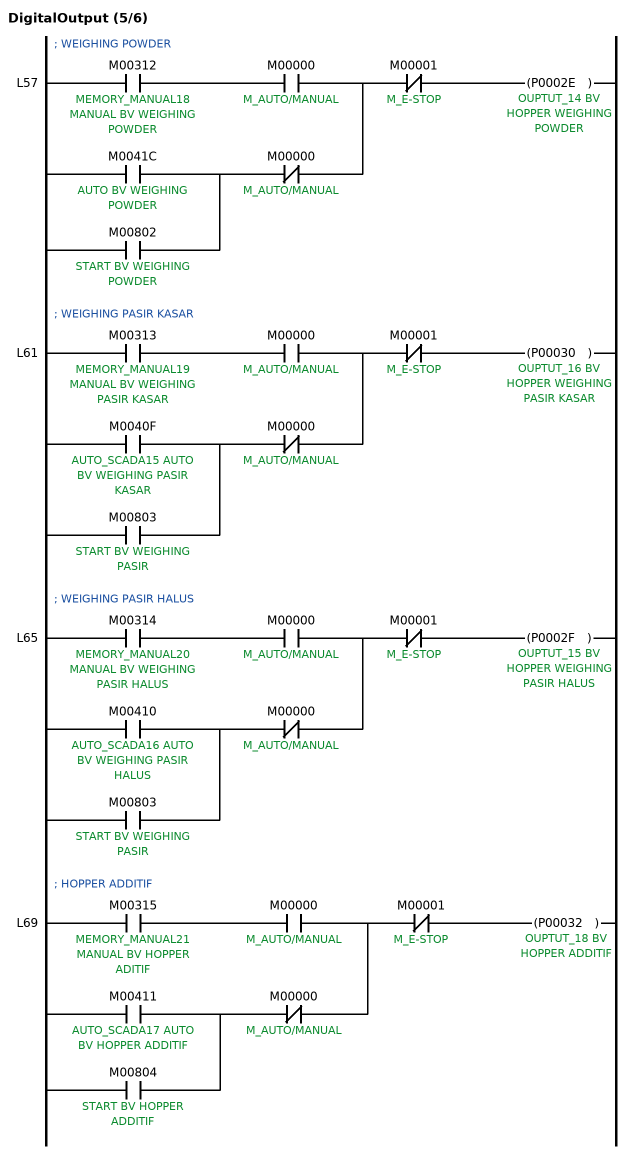
// WEIGHING POWDER
; L57
LOAD      M00312	// MEMORY_MANUAL18 MANUAL BV WEIGHING POWDER 
AND       M00000	// M_AUTO/MANUAL
LOAD      M0041C	// AUTO BV WEIGHING POWDER
OR        M00802	// START BV WEIGHING POWDER 
AND NOT   M00000	// M_AUTO/MANUAL
OR LOAD
AND NOT   M00001	// M_E-STOP
OUT       P0002E	// OUPTUT_14 BV HOPPER WEIGHING POWDER
// WEIGHING PASIR KASAR
; L61
LOAD      M00313	// MEMORY_MANUAL19 MANUAL BV WEIGHING PASIR KASAR 
AND       M00000	// M_AUTO/MANUAL
LOAD      M0040F	// AUTO_SCADA15 AUTO BV WEIGHING PASIR KASAR 
OR        M00803	// START BV WEIGHING PASIR 
AND NOT   M00000	// M_AUTO/MANUAL
OR LOAD
AND NOT   M00001	// M_E-STOP
OUT       P00030	// OUPTUT_16 BV HOPPER WEIGHING PASIR KASAR
// WEIGHING PASIR HALUS
; L65
LOAD      M00314	// MEMORY_MANUAL20 MANUAL BV WEIGHING PASIR HALUS 
AND       M00000	// M_AUTO/MANUAL
LOAD      M00410	// AUTO_SCADA16 AUTO BV WEIGHING PASIR HALUS 
OR        M00803	// START BV WEIGHING PASIR 
AND NOT   M00000	// M_AUTO/MANUAL
OR LOAD
AND NOT   M00001	// M_E-STOP
OUT       P0002F	// OUPTUT_15 BV HOPPER WEIGHING PASIR HALUS
// HOPPER ADDITIF
; L69
LOAD      M00315	// MEMORY_MANUAL21 MANUAL BV HOPPER ADITIF 
AND       M00000	// M_AUTO/MANUAL
LOAD      M00411	// AUTO_SCADA17 AUTO BV HOPPER ADDITIF 
OR        M00804	// START BV HOPPER ADDITIF 
AND NOT   M00000	// M_AUTO/MANUAL
OR LOAD
AND NOT   M00001	// M_E-STOP
OUT       P00032	// OUPTUT_18 BV HOPPER ADDITIF

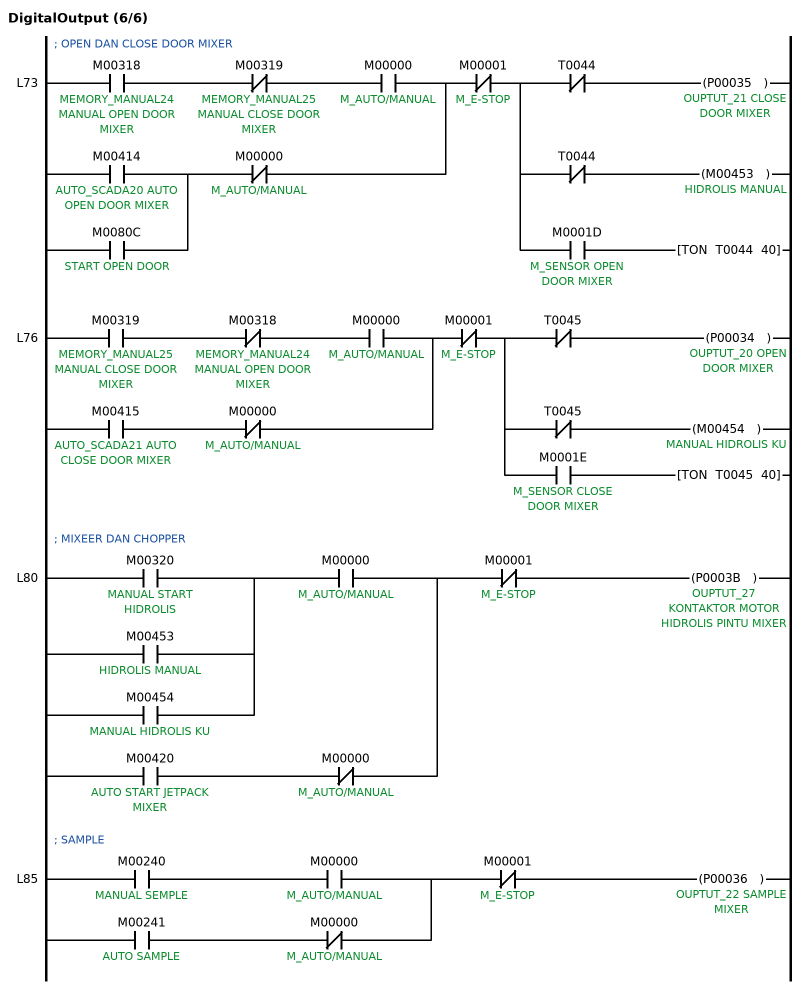
// OPEN DAN CLOSE DOOR MIXER
; L73
LOAD      M00318	// MEMORY_MANUAL24 MANUAL OPEN DOOR MIXER 
AND NOT   M00319	// MEMORY_MANUAL25 MANUAL CLOSE DOOR MIXER 
AND       M00000	// M_AUTO/MANUAL
LOAD      M00414	// AUTO_SCADA20 AUTO OPEN DOOR MIXER 
OR        M0080C	// START OPEN DOOR 
AND NOT   M00000	// M_AUTO/MANUAL
OR LOAD
AND NOT   M00001	// M_E-STOP
MPUSH
AND NOT   T0044
OUT       P00035	// OUPTUT_21 CLOSE DOOR MIXER 
MLOAD
AND NOT   T0044
OUT       M00453	// HIDROLIS MANUAL
MPOP
AND       M0001D	// M_SENSOR OPEN DOOR MIXER 
TON       T0044 40
; L76
LOAD      M00319	// MEMORY_MANUAL25 MANUAL CLOSE DOOR MIXER 
AND NOT   M00318	// MEMORY_MANUAL24 MANUAL OPEN DOOR MIXER 
AND       M00000	// M_AUTO/MANUAL
LOAD      M00415	// AUTO_SCADA21 AUTO CLOSE DOOR MIXER 
AND NOT   M00000	// M_AUTO/MANUAL
OR LOAD
AND NOT   M00001	// M_E-STOP
MPUSH
AND NOT   T0045
OUT       P00034	// OUPTUT_20 OPEN DOOR MIXER 
MLOAD
AND NOT   T0045
OUT       M00454	// MANUAL HIDROLIS KU
MPOP
AND       M0001E	// M_SENSOR CLOSE DOOR MIXER
TON       T0045 40
// MIXEER DAN CHOPPER
; L80
LOAD      M00320	// MANUAL START HIDROLIS
OR        M00453	// HIDROLIS MANUAL
OR        M00454	// MANUAL HIDROLIS KU
AND       M00000	// M_AUTO/MANUAL
LOAD      M00420	// AUTO START JETPACK  MIXER
AND NOT   M00000	// M_AUTO/MANUAL
OR LOAD
AND NOT   M00001	// M_E-STOP
OUT       P0003B	// OUPTUT_27 KONTAKTOR MOTOR HIDROLIS PINTU MIXER
// SAMPLE
; L85
LOAD      M00240	// MANUAL SEMPLE
AND       M00000	// M_AUTO/MANUAL
LOAD      M00241	// AUTO SAMPLE
AND NOT   M00000	// M_AUTO/MANUAL
OR LOAD
AND NOT   M00001	// M_E-STOP
OUT       P00036	// OUPTUT_22 SAMPLE MIXER 

PROGRAM FeedingAdditif (task: Scan Program)

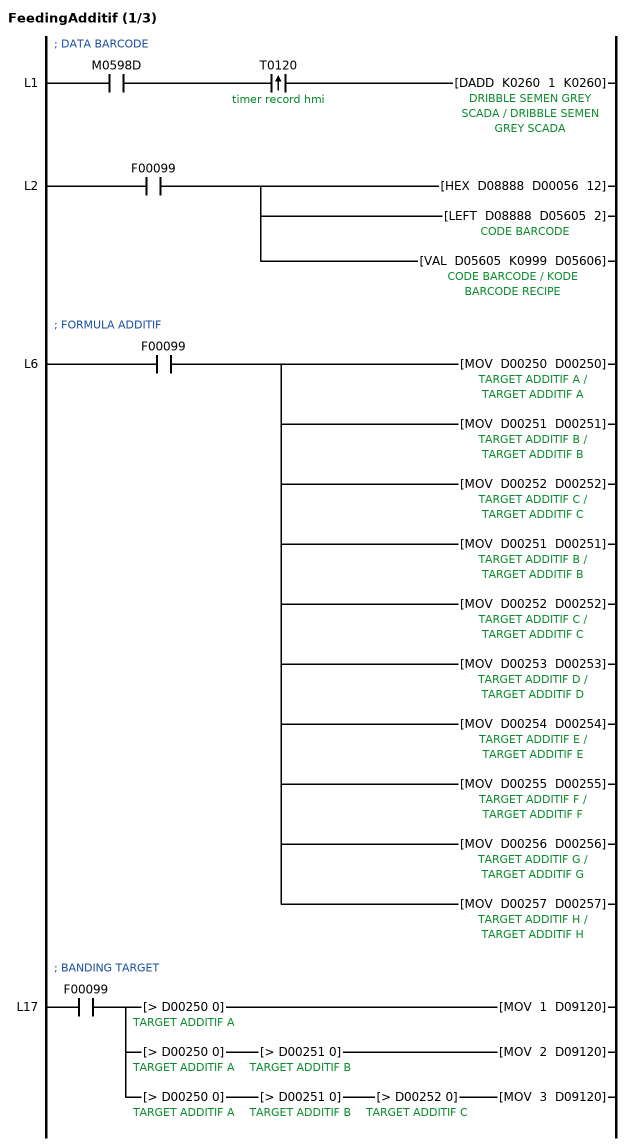
// DATA BARCODE
; L1
LOAD      M0598D
ANDP      T0120	// timer record hmi
DADD      K0260 1 K0260	// DRIBBLE SEMEN GREY SCADA / DRIBBLE SEMEN GREY SCADA
; L2
LOAD      F00099
HEX       D08888 D00056 12
LEFT      D08888 D05605 2	// CODE BARCODE
VAL       D05605 K0999 D05606	// CODE BARCODE / KODE BARCODE RECIPE
// FORMULA ADDITIF
; L6
LOAD      F00099
MOV       D00250 D00250	// TARGET ADDITIF A / TARGET ADDITIF A
MOV       D00251 D00251	// TARGET ADDITIF B / TARGET ADDITIF B
MOV       D00252 D00252	// TARGET ADDITIF C / TARGET ADDITIF C
MOV       D00251 D00251	// TARGET ADDITIF B / TARGET ADDITIF B
MOV       D00252 D00252	// TARGET ADDITIF C / TARGET ADDITIF C
MOV       D00253 D00253	// TARGET ADDITIF D / TARGET ADDITIF D
MOV       D00254 D00254	// TARGET ADDITIF E / TARGET ADDITIF E
MOV       D00255 D00255	// TARGET ADDITIF F / TARGET ADDITIF F
MOV       D00256 D00256	// TARGET ADDITIF G / TARGET ADDITIF G
MOV       D00257 D00257	// TARGET ADDITIF H / TARGET ADDITIF H
// BANDING TARGET
; L17
LOAD      F00099
MPUSH
AND>      D00250 0	// TARGET ADDITIF A
MOV       1 D09120
MLOAD
AND>      D00250 0	// TARGET ADDITIF A
AND>      D00251 0	// TARGET ADDITIF B
MOV       2 D09120
MPOP
AND>      D00250 0	// TARGET ADDITIF A
AND>      D00251 0	// TARGET ADDITIF B
AND>      D00252 0	// TARGET ADDITIF C
MOV       3 D09120

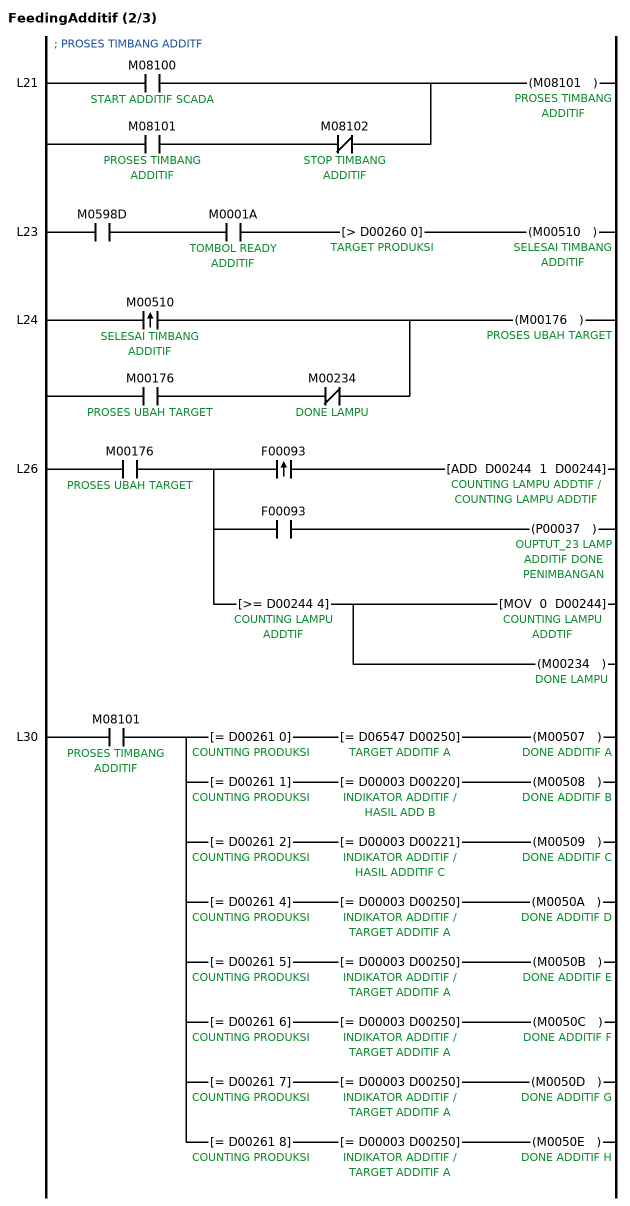
// PROSES TIMBANG ADDITF
; L21
LOAD      M08100	// START ADDITIF SCADA
LOAD      M08101	// PROSES TIMBANG ADDITIF
AND NOT   M08102	// STOP TIMBANG ADDITIF
OR LOAD
OUT       M08101	// PROSES TIMBANG ADDITIF
; L23
LOAD      M0598D
AND       M0001A	// TOMBOL READY ADDITIF
AND>      D00260 0	// TARGET PRODUKSI 
OUT       M00510	// SELESAI TIMBANG  ADDITIF 
; L24
LOADP     M00510	// SELESAI TIMBANG  ADDITIF 
LOAD      M00176	// PROSES UBAH TARGET
AND NOT   M00234	// DONE LAMPU
OR LOAD
OUT       M00176	// PROSES UBAH TARGET
; L26
LOAD      M00176	// PROSES UBAH TARGET
MPUSH
ANDP      F00093
ADD       D00244 1 D00244	// COUNTING LAMPU ADDTIF / COUNTING LAMPU ADDTIF
MLOAD
AND       F00093
OUT       P00037	// OUPTUT_23 LAMP ADDITIF DONE PENIMBANGAN
MPOP
AND>=     D00244 4	// COUNTING LAMPU ADDTIF
MOV       0 D00244	// COUNTING LAMPU ADDTIF
OUT       M00234	// DONE LAMPU
; L30
LOAD      M08101	// PROSES TIMBANG ADDITIF
MPUSH
AND=      D00261 0	// COUNTING PRODUKSI
AND=      D06547 D00250	// TARGET ADDITIF A
OUT       M00507	// DONE ADDITIF A
MLOAD
AND=      D00261 1	// COUNTING PRODUKSI
AND=      D00003 D00220	// INDIKATOR ADDITIF / HASIL ADD B
OUT       M00508	// DONE ADDITIF B
MLOAD
AND=      D00261 2	// COUNTING PRODUKSI
AND=      D00003 D00221	// INDIKATOR ADDITIF / HASIL ADDITIF C
OUT       M00509	// DONE ADDITIF C
MLOAD
AND=      D00261 4	// COUNTING PRODUKSI
AND=      D00003 D00250	// INDIKATOR ADDITIF / TARGET ADDITIF A
OUT       M0050A	// DONE ADDITIF D
MLOAD
AND=      D00261 5	// COUNTING PRODUKSI
AND=      D00003 D00250	// INDIKATOR ADDITIF / TARGET ADDITIF A
OUT       M0050B	// DONE ADDITIF E
MLOAD
AND=      D00261 6	// COUNTING PRODUKSI
AND=      D00003 D00250	// INDIKATOR ADDITIF / TARGET ADDITIF A
OUT       M0050C	// DONE ADDITIF F
MLOAD
AND=      D00261 7	// COUNTING PRODUKSI
AND=      D00003 D00250	// INDIKATOR ADDITIF / TARGET ADDITIF A
OUT       M0050D	// DONE ADDITIF G
MPOP
AND=      D00261 8	// COUNTING PRODUKSI
AND=      D00003 D00250	// INDIKATOR ADDITIF / TARGET ADDITIF A
OUT       M0050E	// DONE ADDITIF H

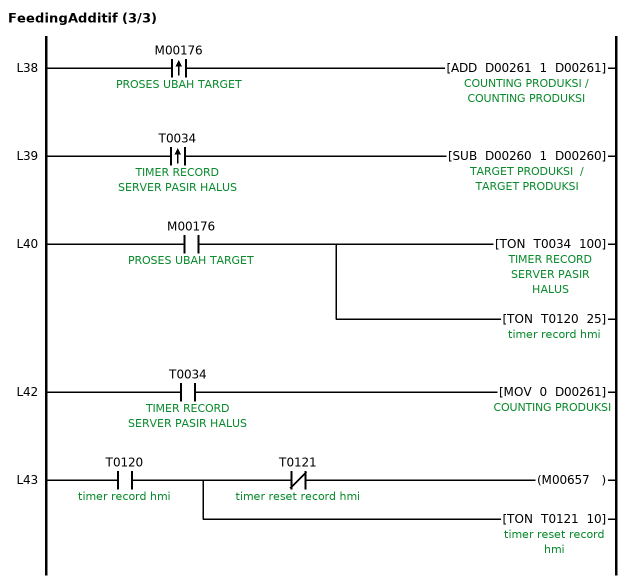
; L38
LOADP     M00176	// PROSES UBAH TARGET
ADD       D00261 1 D00261	// COUNTING PRODUKSI / COUNTING PRODUKSI
; L39
LOADP     T0034	// TIMER RECORD SERVER PASIR HALUS
SUB       D00260 1 D00260	// TARGET PRODUKSI  / TARGET PRODUKSI 
; L40
LOAD      M00176	// PROSES UBAH TARGET
TON       T0034 100	// TIMER RECORD SERVER PASIR HALUS
TON       T0120 25	// timer record hmi
; L42
LOAD      T0034	// TIMER RECORD SERVER PASIR HALUS
MOV       0 D00261	// COUNTING PRODUKSI
; L43
LOAD      T0120	// timer record hmi
MPUSH
AND NOT   T0121	// timer reset record hmi
OUT       M00657
MPOP
TON       T0121 10	// timer reset record hmi

PROGRAM ProsesFeedingMaterial (task: Scan Program)

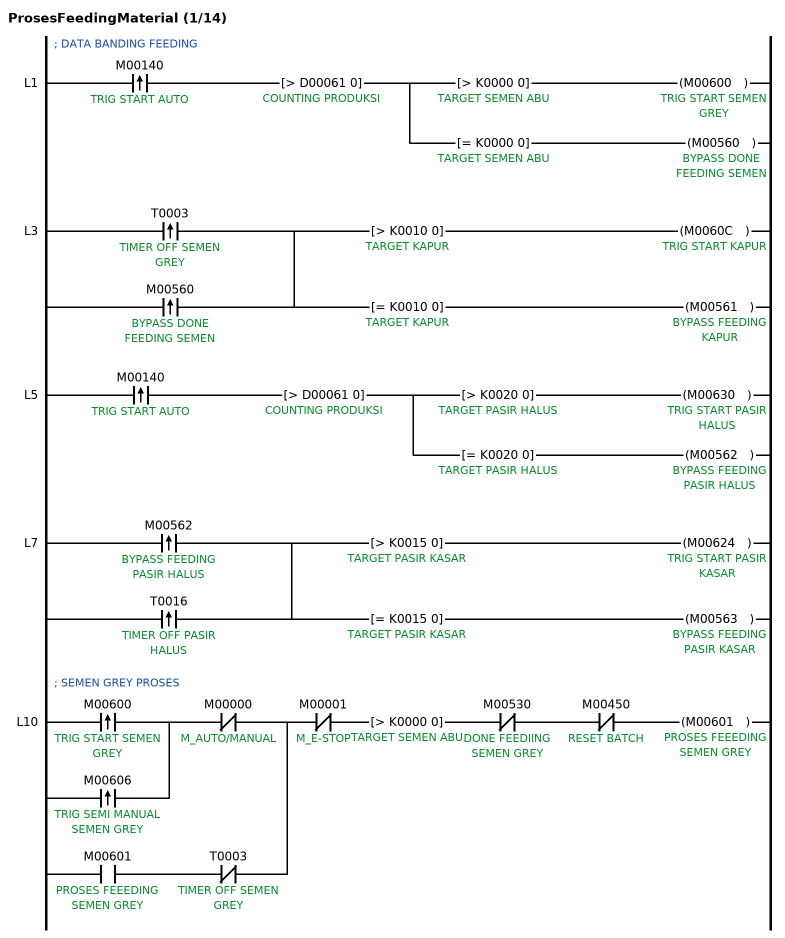
// DATA BANDING FEEDING
; L1
LOADP     M00140	// TRIG START AUTO
AND>      D00061 0	// COUNTING PRODUKSI
MPUSH
AND>      K0000 0	// TARGET SEMEN ABU 
OUT       M00600	// TRIG START SEMEN GREY 
MPOP
AND=      K0000 0	// TARGET SEMEN ABU 
OUT       M00560	// BYPASS DONE FEEDING SEMEN
; L3
LOADP     T0003	// TIMER OFF SEMEN GREY 
ORP       M00560	// BYPASS DONE FEEDING SEMEN
MPUSH
AND>      K0010 0	// TARGET KAPUR 
OUT       M0060C	// TRIG START KAPUR
MPOP
AND=      K0010 0	// TARGET KAPUR 
OUT       M00561	// BYPASS FEEDING KAPUR
; L5
LOADP     M00140	// TRIG START AUTO
AND>      D00061 0	// COUNTING PRODUKSI
MPUSH
AND>      K0020 0	// TARGET PASIR HALUS 
OUT       M00630	// TRIG START PASIR HALUS
MPOP
AND=      K0020 0	// TARGET PASIR HALUS 
OUT       M00562	// BYPASS FEEDING PASIR HALUS
; L7
LOADP     M00562	// BYPASS FEEDING PASIR HALUS
ORP       T0016	// TIMER OFF PASIR HALUS 
MPUSH
AND>      K0015 0	// TARGET PASIR KASAR
OUT       M00624	// TRIG START PASIR KASAR
MPOP
AND=      K0015 0	// TARGET PASIR KASAR
OUT       M00563	// BYPASS FEEDING PASIR KASAR
// SEMEN GREY PROSES
; L10
LOADP     M00600	// TRIG START SEMEN GREY 
ORP       M00606	// TRIG SEMI MANUAL SEMEN GREY 
AND NOT   M00000	// M_AUTO/MANUAL
LOAD      M00601	// PROSES FEEEDING SEMEN GREY
AND NOT   T0003	// TIMER OFF SEMEN GREY 
OR LOAD
AND NOT   M00001	// M_E-STOP
AND>      K0000 0	// TARGET SEMEN ABU 
AND NOT   M00530	// DONE FEEDIING SEMEN GREY 
AND NOT   M00450	// RESET BATCH
OUT       M00601	// PROSES FEEEDING SEMEN GREY

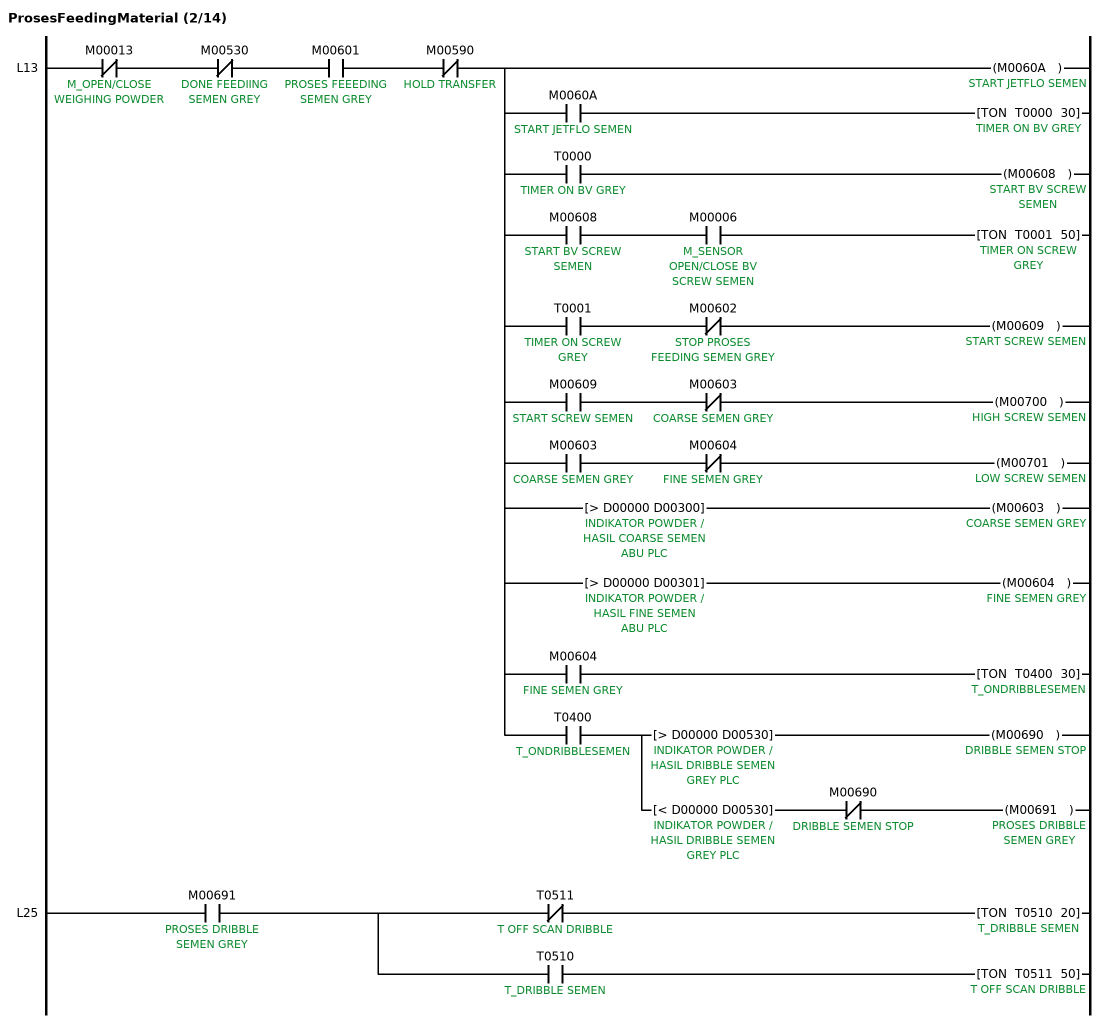
; L13
LOAD NOT  M00013	// M_OPEN/CLOSE WEIGHING POWDER
AND NOT   M00530	// DONE FEEDIING SEMEN GREY 
AND       M00601	// PROSES FEEEDING SEMEN GREY
AND NOT   M00590	// HOLD TRANSFER
OUT       M0060A	// START JETFLO SEMEN
MPUSH
AND       M0060A	// START JETFLO SEMEN
TON       T0000 30	// TIMER ON BV GREY
MLOAD
AND       T0000	// TIMER ON BV GREY
OUT       M00608	// START BV SCREW SEMEN 
MLOAD
AND       M00608	// START BV SCREW SEMEN 
AND       M00006	// M_SENSOR OPEN/CLOSE BV SCREW SEMEN
TON       T0001 50	// TIMER ON SCREW GREY 
MLOAD
AND       T0001	// TIMER ON SCREW GREY 
AND NOT   M00602	// STOP PROSES FEEDING SEMEN GREY 
OUT       M00609	// START SCREW SEMEN
MLOAD
AND       M00609	// START SCREW SEMEN
AND NOT   M00603	// COARSE SEMEN GREY
OUT       M00700	// HIGH SCREW SEMEN
MLOAD
AND       M00603	// COARSE SEMEN GREY
AND NOT   M00604	// FINE SEMEN GREY
OUT       M00701	// LOW SCREW SEMEN
MLOAD
AND>      D00000 D00300	// INDIKATOR POWDER / HASIL COARSE SEMEN ABU PLC
OUT       M00603	// COARSE SEMEN GREY
MLOAD
AND>      D00000 D00301	// INDIKATOR POWDER / HASIL FINE SEMEN ABU PLC
OUT       M00604	// FINE SEMEN GREY
MLOAD
AND       M00604	// FINE SEMEN GREY
TON       T0400 30	// T_ONDRIBBLESEMEN
MPOP
AND       T0400	// T_ONDRIBBLESEMEN
MPUSH
AND>      D00000 D00530	// INDIKATOR POWDER / HASIL DRIBBLE SEMEN GREY PLC
OUT       M00690	// DRIBBLE SEMEN STOP
MPOP
AND<      D00000 D00530	// INDIKATOR POWDER / HASIL DRIBBLE SEMEN GREY PLC
AND NOT   M00690	// DRIBBLE SEMEN STOP
OUT       M00691	// PROSES DRIBBLE SEMEN GREY
; L25
LOAD      M00691	// PROSES DRIBBLE SEMEN GREY
MPUSH
AND NOT   T0511	// T OFF SCAN DRIBBLE
TON       T0510 20	// T_DRIBBLE SEMEN
MPOP
AND       T0510	// T_DRIBBLE SEMEN
TON       T0511 50	// T OFF SCAN DRIBBLE

